FUNCTION_BLOCK "FB_PressDemoAuto"
{ S7_Optimized_Access := 'TRUE' }
VERSION : 0.1
VAR_INPUT
    Run : Bool;
    Reset : Bool;
    OwnerIndex : DInt;
    Delta : Time;
    TransferSettleTime : Time;
    PartQuality : Bool;
    RequireTwoHandStart : Bool;
    SourcePath : String[80];
    PartPresent : Bool;
    AirPressureOk : Bool;
    TwoHandHeld : Bool;
    StartPulse : Bool;
    PressSettleTime : Time;
END_VAR
VAR_IN_OUT
    PressRam {ExternalAccessible := 'False'; ExternalVisible := 'False'; ExternalWritable := 'False'} : "FB_CylinderCM";
    Door {ExternalAccessible := 'False'; ExternalVisible := 'False'; ExternalWritable := 'False'} : "FB_CylinderCM";
    PartSlide {ExternalAccessible := 'False'; ExternalVisible := 'False'; ExternalWritable := 'False'} : "FB_CylinderCM";
    Core {ExternalAccessible := 'False'; ExternalVisible := 'False'; ExternalWritable := 'False'} : "FRK_Core";
    Unit {ExternalAccessible := 'False'; ExternalVisible := 'False'; ExternalWritable := 'False'} : "FRK_Unit";
    Status {ExternalAccessible := 'False'; ExternalVisible := 'False'; ExternalWritable := 'False'} : "ST_ModuleStatus";
    Part {ExternalAccessible := 'False'; ExternalVisible := 'False'; ExternalWritable := 'False'} : "ST_PartContext";
    AlarmLog {ExternalAccessible := 'False'; ExternalVisible := 'False'; ExternalWritable := 'False'} : "FRK_AlarmLog";
END_VAR
VAR_OUTPUT
END_VAR
VAR
    Seq {ExternalWritable := 'False'} : "FRK_SequenceCtx";
    Row1 {ExternalWritable := 'False'} : "FRK_SequenceRow";
    Row2 {ExternalWritable := 'False'} : "FRK_SequenceRow";
    Row3 {ExternalWritable := 'False'} : "FRK_SequenceRow";
    Row4 {ExternalWritable := 'False'} : "FRK_SequenceRow";
    Row5 {ExternalWritable := 'False'} : "FRK_SequenceRow";
    Row6 {ExternalWritable := 'False'} : "FRK_SequenceRow";
    Row7 {ExternalWritable := 'False'} : "FRK_SequenceRow";
    Row8 {ExternalWritable := 'False'} : "FRK_SequenceRow";
    Row9 {ExternalWritable := 'False'} : "FRK_SequenceRow";
    Row10 {ExternalWritable := 'False'} : "FRK_SequenceRow";
    Row11 {ExternalWritable := 'False'} : "FRK_SequenceRow";
    Row12 {ExternalWritable := 'False'} : "FRK_SequenceRow";
    Row13 {ExternalWritable := 'False'} : "FRK_SequenceRow";
    Row14 {ExternalWritable := 'False'} : "FRK_SequenceRow";
    Row15 {ExternalWritable := 'False'} : "FRK_SequenceRow";
    Row16 {ExternalWritable := 'False'} : "FRK_SequenceRow";
    At0 {ExternalAccessible := 'False'; ExternalVisible := 'False'; ExternalWritable := 'False'} : Bool;
    At100 {ExternalAccessible := 'False'; ExternalVisible := 'False'; ExternalWritable := 'False'} : Bool;
    At110 {ExternalAccessible := 'False'; ExternalVisible := 'False'; ExternalWritable := 'False'} : Bool;
    At130 {ExternalAccessible := 'False'; ExternalVisible := 'False'; ExternalWritable := 'False'} : Bool;
    At150 {ExternalAccessible := 'False'; ExternalVisible := 'False'; ExternalWritable := 'False'} : Bool;
    At170 {ExternalAccessible := 'False'; ExternalVisible := 'False'; ExternalWritable := 'False'} : Bool;
    At180 {ExternalAccessible := 'False'; ExternalVisible := 'False'; ExternalWritable := 'False'} : Bool;
    At185 {ExternalAccessible := 'False'; ExternalVisible := 'False'; ExternalWritable := 'False'} : Bool;
    At190 {ExternalAccessible := 'False'; ExternalVisible := 'False'; ExternalWritable := 'False'} : Bool;
    At200 {ExternalAccessible := 'False'; ExternalVisible := 'False'; ExternalWritable := 'False'} : Bool;
    At210 {ExternalAccessible := 'False'; ExternalVisible := 'False'; ExternalWritable := 'False'} : Bool;
    At215 {ExternalAccessible := 'False'; ExternalVisible := 'False'; ExternalWritable := 'False'} : Bool;
    At220 {ExternalAccessible := 'False'; ExternalVisible := 'False'; ExternalWritable := 'False'} : Bool;
    At230 {ExternalAccessible := 'False'; ExternalVisible := 'False'; ExternalWritable := 'False'} : Bool;
    At240 {ExternalAccessible := 'False'; ExternalVisible := 'False'; ExternalWritable := 'False'} : Bool;
    At999 {ExternalAccessible := 'False'; ExternalVisible := 'False'; ExternalWritable := 'False'} : Bool;
    Ready1 {ExternalAccessible := 'False'; ExternalVisible := 'False'; ExternalWritable := 'False'} : Bool;
    Ready2 {ExternalAccessible := 'False'; ExternalVisible := 'False'; ExternalWritable := 'False'} : Bool;
    Ready3 {ExternalAccessible := 'False'; ExternalVisible := 'False'; ExternalWritable := 'False'} : Bool;
    Ready4 {ExternalAccessible := 'False'; ExternalVisible := 'False'; ExternalWritable := 'False'} : Bool;
    Ready5 {ExternalAccessible := 'False'; ExternalVisible := 'False'; ExternalWritable := 'False'} : Bool;
    Advance {ExternalAccessible := 'False'; ExternalVisible := 'False'; ExternalWritable := 'False'} : Bool;
    Cycle {ExternalAccessible := 'False'; ExternalVisible := 'False'; ExternalWritable := 'False'} : "ST_PressDemoCycle";
    LoadPosition {ExternalAccessible := 'False'; ExternalVisible := 'False'; ExternalWritable := 'False'} : "FB_PressDemoLoadPosition";
    LoadDone {ExternalAccessible := 'False'; ExternalVisible := 'False'; ExternalWritable := 'False'} : Bool;
    LoadActive {ExternalAccessible := 'False'; ExternalVisible := 'False'; ExternalWritable := 'False'} : Bool;
END_VAR
BEGIN
    "FRK_SeqBegin"(Run := #Run, Reset := #Reset, OwnerIndex := #OwnerIndex, ChainIndex := 1, BranchIndex := 0, ViewOffset := 0, ViewDepth := 0, Delta := #Delta, Seq := #Seq);
    "FRK_SeqStart"(Seq := #Seq, StartPulse := #StartPulse);
    "F_PressDemoReset"(Seq := #Seq, Cycle := #Cycle);
    #LoadActive := "FRK_SeqSubActive"(Seq := #Seq, Run := #Run, StepNo := 240);
    #LoadDone := "F_PressDemoLoadPosition"(Target := #LoadPosition, Run := #LoadActive, Reset := #Seq.Restart OR #Seq.Rearm, OwnerIndex := #OwnerIndex, Delta := #Delta, PressRam := #PressRam, Door := #Door, PartSlide := #PartSlide);
    "F_CylinderSequenceLease"(Seq := #Seq, Target := #PressRam);
    "F_CylinderSequenceLease"(Seq := #Seq, Target := #Door);
    "F_CylinderSequenceLease"(Seq := #Seq, Target := #PartSlide);
    "FRK_SeqOwnerStatus"(Seq := #Seq, Core := #Core, Status := #Status);
    "FRK_SeqSubStatus"(Seq := #Seq, Child := #LoadPosition.Seq);
    CASE #Seq.ScanStep OF
        0:
            IF #Seq.Running AND NOT #Seq.Error THEN
                "FRK_SeqStep"(StepNo := 0, StepName := 'project.step.pressAutoInitialize', AwaitingLabel := '', AwaitsPath := '', TimeClass := 0, ExpectedTime := #Seq.NoTimeGuard, Seq := #Seq, Row := #Row1);
                "FRK_SeqReady"(Seq := #Seq, Ok1 := TRUE, Ok2 := TRUE, Ok3 := TRUE, Ok4 := TRUE, Ok5 := TRUE);
                "FRK_SeqRoute"(Seq := #Seq, OnAdvance := 100, OnJump1 := -1);
            END_IF;
        100:
            IF #Seq.Running AND NOT #Seq.Error THEN
                "FRK_SeqStep"(StepNo := 100, StepName := 'project.step.pressAwaitTwoHand', AwaitingLabel := '', AwaitsPath := '', TimeClass := 3, ExpectedTime := #Seq.NoTimeGuard, Seq := #Seq, Row := #Row2);
                #Ready5 := "F_PressDemoAwaitCycle"(Seq := #Seq, Cycle := #Cycle, Core := #Core, Unit := #Unit, Status := #Status, Part := #Part, AlarmLog := #AlarmLog, PartPresent := #PartPresent, PartQuality := #PartQuality, AirPressureOk := #AirPressureOk, RequireTwoHandStart := #RequireTwoHandStart);
                "FRK_SeqReady"(Seq := #Seq, Ok1 := #Ready5, Ok2 := TRUE, Ok3 := TRUE, Ok4 := TRUE, Ok5 := TRUE);
                "FRK_SeqRoute"(Seq := #Seq, OnAdvance := 110, OnJump1 := -1);
            END_IF;
        110:
            IF #Seq.Running AND NOT #Seq.Error THEN
                "FRK_SeqStep"(StepNo := 110, StepName := 'project.step.pressRamUp', AwaitingLabel := 'PressRam.RETRACT', AwaitsPath := #PressRam.Status.Name, TimeClass := 0, ExpectedTime := #Seq.NoTimeGuard, Seq := #Seq, Row := #Row3);
                #Ready1 := "F_CylinderRetract"(Seq := #Seq, Target := #PressRam);
                "FRK_SeqReady"(Seq := #Seq, Ok1 := #Ready1, Ok2 := TRUE, Ok3 := TRUE, Ok4 := TRUE, Ok5 := TRUE);
                "FRK_SeqRoute"(Seq := #Seq, OnAdvance := 130, OnJump1 := -1);
            END_IF;
        130:
            IF #Seq.Running AND NOT #Seq.Error THEN
                "FRK_SeqStep"(StepNo := 130, StepName := 'project.step.pressDoorOpen', AwaitingLabel := 'Door.RETRACT', AwaitsPath := #Door.Status.Name, TimeClass := 0, ExpectedTime := #Seq.NoTimeGuard, Seq := #Seq, Row := #Row4);
                #Ready1 := "F_CylinderRetract"(Seq := #Seq, Target := #Door);
                "FRK_SeqReady"(Seq := #Seq, Ok1 := #Ready1, Ok2 := TRUE, Ok3 := TRUE, Ok4 := TRUE, Ok5 := TRUE);
                "FRK_SeqRoute"(Seq := #Seq, OnAdvance := 150, OnJump1 := -1);
            END_IF;
        150:
            IF #Seq.Running AND NOT #Seq.Error THEN
                "FRK_SeqStep"(StepNo := 150, StepName := 'project.step.pressSlideInside', AwaitingLabel := 'PartSlide.EXTEND', AwaitsPath := #PartSlide.Status.Name, TimeClass := 0, ExpectedTime := #Seq.NoTimeGuard, Seq := #Seq, Row := #Row5);
                #Ready1 := "F_CylinderExtend"(Seq := #Seq, Target := #PartSlide);
                "F_PressDemoStarted"(Seq := #Seq, Unit := #Unit, Status := #Status, Part := #Part, AlarmLog := #AlarmLog);
                "FRK_SeqReady"(Seq := #Seq, Ok1 := #Ready1, Ok2 := TRUE, Ok3 := TRUE, Ok4 := TRUE, Ok5 := TRUE);
                "FRK_SeqRoute"(Seq := #Seq, OnAdvance := 170, OnJump1 := -1);
            END_IF;
        170:
            IF #Seq.Running AND NOT #Seq.Error THEN
                "FRK_SeqStep"(StepNo := 170, StepName := 'project.step.pressTransferSettle', AwaitingLabel := '', AwaitsPath := '', TimeClass := 0, ExpectedTime := #TransferSettleTime, Seq := #Seq, Row := #Row6);
                #Ready1 := "FRK_SeqDelay"(Seq := #Seq, PT := #TransferSettleTime, Delta := #Delta, Permit := TRUE);
                "FRK_SeqReady"(Seq := #Seq, Ok1 := #Ready1, Ok2 := TRUE, Ok3 := TRUE, Ok4 := TRUE, Ok5 := TRUE);
                "FRK_SeqRoute"(Seq := #Seq, OnAdvance := 180, OnJump1 := -1);
            END_IF;
        180:
            IF #Seq.Running AND NOT #Seq.Error THEN
                "FRK_SeqStep"(StepNo := 180, StepName := 'project.step.pressDoorClose', AwaitingLabel := 'Door.EXTEND', AwaitsPath := #Door.Status.Name, TimeClass := 0, ExpectedTime := #Seq.NoTimeGuard, Seq := #Seq, Row := #Row7);
                #Ready1 := "F_CylinderExtend"(Seq := #Seq, Target := #Door);
                "F_PressDemoDoorClose"(Seq := #Seq, Closed := #Ready1, TwoHandHeld := #TwoHandHeld, RequireTwoHandStart := #RequireTwoHandStart, SourcePath := #SourcePath, AlarmLog := #AlarmLog);
                "FRK_SeqRoute"(Seq := #Seq, OnAdvance := 200, OnJump1 := 185);
            END_IF;
        185:
            IF #Seq.Running AND NOT #Seq.Error THEN
                "FRK_SeqStep"(StepNo := 185, StepName := 'project.step.pressDoorReopen', AwaitingLabel := 'Door.RETRACT', AwaitsPath := #Door.Status.Name, TimeClass := 0, ExpectedTime := #Seq.NoTimeGuard, Seq := #Seq, Row := #Row8);
                #Ready1 := "F_CylinderRetract"(Seq := #Seq, Target := #Door);
                "FRK_SeqReady"(Seq := #Seq, Ok1 := #Ready1, Ok2 := TRUE, Ok3 := TRUE, Ok4 := TRUE, Ok5 := TRUE);
                "FRK_SeqRoute"(Seq := #Seq, OnAdvance := 190, OnJump1 := -1);
            END_IF;
        190:
            IF #Seq.Running AND NOT #Seq.Error THEN
                "FRK_SeqStep"(StepNo := 190, StepName := 'project.step.pressSlideOutsideAfterAbort', AwaitingLabel := 'PartSlide.RETRACT', AwaitsPath := #PartSlide.Status.Name, TimeClass := 0, ExpectedTime := #Seq.NoTimeGuard, Seq := #Seq, Row := #Row9);
                #Ready1 := "F_CylinderRetract"(Seq := #Seq, Target := #PartSlide);
                "F_PressDemoClearStart"(Seq := #Seq, Complete := #Ready1);
                "FRK_SeqReady"(Seq := #Seq, Ok1 := #Ready1, Ok2 := TRUE, Ok3 := TRUE, Ok4 := TRUE, Ok5 := TRUE);
                "FRK_SeqRoute"(Seq := #Seq, OnAdvance := 100, OnJump1 := -1);
            END_IF;
        200:
            IF #Seq.Running AND NOT #Seq.Error THEN
                "FRK_SeqStep"(StepNo := 200, StepName := 'project.step.pressRamDown', AwaitingLabel := 'PressRam.EXTEND', AwaitsPath := #PressRam.Status.Name, TimeClass := 0, ExpectedTime := #Seq.NoTimeGuard, Seq := #Seq, Row := #Row10);
                #Ready1 := "F_CylinderExtendHandled"(Seq := #Seq, Target := #PressRam);
                "F_PressDemoRamResult"(Seq := #Seq, Reached := #Ready1, Cycle := #Cycle, AlarmLog := #AlarmLog);
                "FRK_SeqRoute"(Seq := #Seq, OnAdvance := 220, OnJump1 := 210);
            END_IF;
        210:
            IF #Seq.Running AND NOT #Seq.Error THEN
                "FRK_SeqStep"(StepNo := 210, StepName := 'project.step.pressNotReachedConfirm', AwaitingLabel := '', AwaitsPath := '', TimeClass := 3, ExpectedTime := #Seq.NoTimeGuard, Seq := #Seq, Row := #Row11);
                #Ready5 := "F_PressDemoConfirmScrap"(Seq := #Seq, SourcePath := #SourcePath, AlarmLog := #AlarmLog);
                "FRK_SeqReady"(Seq := #Seq, Ok1 := #Ready5, Ok2 := TRUE, Ok3 := TRUE, Ok4 := TRUE, Ok5 := TRUE);
                "FRK_SeqRoute"(Seq := #Seq, OnAdvance := 215, OnJump1 := -1);
            END_IF;
        215:
            IF #Seq.Running AND NOT #Seq.Error THEN
                "FRK_SeqStep"(StepNo := 215, StepName := 'project.step.pressScrapPart', AwaitingLabel := '', AwaitsPath := '', TimeClass := 0, ExpectedTime := #Seq.NoTimeGuard, Seq := #Seq, Row := #Row12);
                #Ready5 := "F_PressDemoScrap"(Seq := #Seq, Cycle := #Cycle, Core := #Core, Unit := #Unit, Status := #Status, Part := #Part, AlarmLog := #AlarmLog);
                "FRK_SeqReady"(Seq := #Seq, Ok1 := #Ready5, Ok2 := TRUE, Ok3 := TRUE, Ok4 := TRUE, Ok5 := TRUE);
                "FRK_SeqRoute"(Seq := #Seq, OnAdvance := 240, OnJump1 := -1);
            END_IF;
        220:
            IF #Seq.Running AND NOT #Seq.Error THEN
                "FRK_SeqStep"(StepNo := 220, StepName := 'project.step.pressDwell', AwaitingLabel := '', AwaitsPath := '', TimeClass := 0, ExpectedTime := #Seq.NoTimeGuard, Seq := #Seq, Row := #Row13);
                #Ready5 := "F_PressDemoDwell"(Seq := #Seq, TwoHandHeld := #TwoHandHeld, RequireTwoHandStart := #RequireTwoHandStart, PT := #PressSettleTime, Delta := #Delta, PressRam := #PressRam);
                "FRK_SeqReady"(Seq := #Seq, Ok1 := #Ready5, Ok2 := TRUE, Ok3 := TRUE, Ok4 := TRUE, Ok5 := TRUE);
                "FRK_SeqRoute"(Seq := #Seq, OnAdvance := 230, OnJump1 := -1);
            END_IF;
        230:
            IF #Seq.Running AND NOT #Seq.Error THEN
                "FRK_SeqStep"(StepNo := 230, StepName := 'project.step.pressRecordResult', AwaitingLabel := '', AwaitsPath := '', TimeClass := 0, ExpectedTime := #Seq.NoTimeGuard, Seq := #Seq, Row := #Row14);
                #Ready5 := "F_PressDemoRecord"(Seq := #Seq, Dwell := #PressSettleTime, Core := #Core, Status := #Status, Part := #Part);
                "FRK_SeqReady"(Seq := #Seq, Ok1 := #Ready5, Ok2 := TRUE, Ok3 := TRUE, Ok4 := TRUE, Ok5 := TRUE);
                "FRK_SeqRoute"(Seq := #Seq, OnAdvance := 240, OnJump1 := -1);
            END_IF;
        240:
            IF #Seq.Running AND NOT #Seq.Error THEN
                "FRK_SeqStep"(StepNo := 240, StepName := 'project.step.pressReturnToLoad', AwaitingLabel := 'project.condition.LoadDone', AwaitsPath := '', TimeClass := 0, ExpectedTime := #Seq.NoTimeGuard, Seq := #Seq, Row := #Row15);
                #Ready1 := "FRK_SeqAwait"(Seq := #Seq, Label := 'project.condition.LoadDone', Ok := #LoadDone);
                "FRK_SeqReady"(Seq := #Seq, Ok1 := #Ready1, Ok2 := TRUE, Ok3 := TRUE, Ok4 := TRUE, Ok5 := TRUE);
                "FRK_SeqRoute"(Seq := #Seq, OnAdvance := 999, OnJump1 := -1);
            END_IF;
        999:
            IF #Seq.Running AND NOT #Seq.Error THEN
                "FRK_SeqStep"(StepNo := 999, StepName := 'project.step.pressAutoComplete', AwaitingLabel := '', AwaitsPath := '', TimeClass := 0, ExpectedTime := #Seq.NoTimeGuard, Seq := #Seq, Row := #Row16);
                #Ready5 := "F_PressDemoCycleEnd"(Seq := #Seq, Cycle := #Cycle, Core := #Core, Unit := #Unit, Status := #Status, Part := #Part, AlarmLog := #AlarmLog);
                "FRK_SeqReady"(Seq := #Seq, Ok1 := #Ready5, Ok2 := TRUE, Ok3 := TRUE, Ok4 := TRUE, Ok5 := TRUE);
                "FRK_SeqRoute"(Seq := #Seq, OnAdvance := 100, OnJump1 := -1);
            END_IF;
        ELSE
            #Seq.Error := TRUE;
            #Seq.ErrorDiagnostic.ReasonCode := 10001;
            #Seq.ErrorDiagnostic.Description := WSTRING#'project.sequence.invalidStep';
    END_CASE;
    "F_CylinderSequenceLease"(Seq := #Seq, Target := #PressRam);
    "F_CylinderSequenceLease"(Seq := #Seq, Target := #Door);
    "F_CylinderSequenceLease"(Seq := #Seq, Target := #PartSlide);
    "FRK_SeqOwnerStatus"(Seq := #Seq, Core := #Core, Status := #Status);
    "FRK_SeqSubStatus"(Seq := #Seq, Child := #LoadPosition.Seq);
END_FUNCTION_BLOCK
